INTERFACE I_Lidar

METHOD Start
END_METHOD

METHOD Stop
END_METHOD

METHOD TryGetScan : BOOL
VAR_INPUT
	scan : REFERENCE TO LaserScan;
END_VAR
END_METHOD

PROPERTY IsRunning : BOOL
GET
END_GET
END_PROPERTY

PROPERTY Error : HardwareError
GET
END_GET
END_PROPERTY

END_INTERFACE

(* stored: Version 1.1.0.1, ProductVersion 3.1.4026.12
   Itf I_Lidar: Id {0d3fe80b-2d66-5794-8f3c-920f32f2296a}
   Method Start: Id {30df7c52-44c0-5d09-be3c-bb9f3e415b7c}
   Method Stop: Id {c74b11f4-71d5-5075-aed5-7395c3032838}
   Method TryGetScan: Id {54ada5e3-844e-52e0-8673-86e30d7c2b37}
   Property IsRunning: Id {54244f47-69ad-597a-ba0e-218a4cb7f82b}
   Get Get: Id {77158aad-602f-5432-8583-c402edf26d8e}
   Property Error: Id {ecf4da05-9385-578f-8431-c111a3eb0b2f}
   Get Get: Id {91eb81ce-d6d6-5fcf-9e61-fd06912f140c} *)
